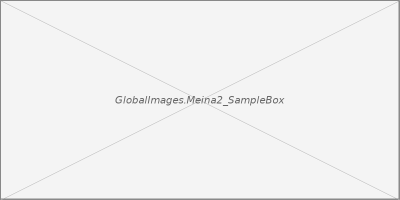
VISUALIZATION V_NCIMeina2_SampleBox  // 400x200
    RoundedRectangle (0,0 400x200)
    Image (0,0 400x200), image: GlobalImages.Meina2_SampleBox
END_VISUALIZATION

(* stored: Version 1.1.0.1, ProductVersion 3.1.4024.15
   Visu V_NCIMeina2_SampleBox: Id {e8acfcc3-d99b-43cb-8296-6fc5c316cb90} *)
